(* IEC 61131-3 sources: s7-to-codesys/src/DUTs/S7Compat, 2 files *)

(* ---- ST_S5Counter.dut.st ---- *)
// Назначение: состояние счётчика S5 (слово счётчика C n S7-300/400) для кода, сконвертированного s7conv из
//             STL: CU, CD, установка S, сброс R, разрешение FR, опрос A C, L C, LC C. Значение 0…999; у
//             каждой инструкции, работающей по фронту RLO, своя память фронта. Состояния лежат в
//             генерируемом GVL_S5Counters (массив aCounter, индекс — номер счётчика).
// Автор:      kr0nsch
// Версия:     1.2.0
// Документ:   docs/MAPPING_STL.md, правило s5.counter
TYPE ST_S5Counter :
STRUCT
    iValue : INT;       // значение счётчика, 0…999
    xRloUp : BOOL;      // RLO последней инструкции CU — память фронта
    xRloDown : BOOL;    // RLO последней инструкции CD — память фронта
    xRloSet : BOOL;     // RLO последней инструкции S — память фронта
    xRloFree : BOOL;    // RLO последней инструкции FR — память фронта разрешения
END_STRUCT
END_TYPE

(* ---- ST_S5Timer.dut.st ---- *)
// Назначение: состояние таймера S5 (слово таймера T n S7-300/400) для кода, сконвертированного s7conv из STL:
//             пуск SP, SE, SD, SS, SF, разрешение FR, сброс R, опрос A T, L T, LC T. В S7 таймер — глобальный
//             объект CPU, поэтому состояния лежат в генерируемом GVL_S5Timers (массив aTimer, индекс — номер
//             таймера), а инструкции — функции F_S5* с VAR_IN_OUT. Время — F_S7Now(): в работе TIME(), в
//             тестах — моделируемые часы GVL_S7Clock. Остаток пересчитывается при каждом обращении к таймеру
//             (в S7 его уменьшает часовой процесс CPU асинхронно циклу).
// Автор:      kr0nsch
// Версия:     1.2.0
// Документ:   docs/MAPPING_STL.md, правило s5.timebase; docs/ASSUMPTIONS.md, записи L13–L16
TYPE ST_S5Timer :
STRUCT
    xRunning : BOOL;    // таймер идёт
    xQ : BOOL;          // состояние таймера (опрос A T n)
    xRloStart : BOOL;   // RLO последней инструкции пуска — память фронта пуска (FR её сбрасывает)
    xRloFree : BOOL;    // RLO последней инструкции FR — память фронта разрешения
    xQAtEnd : BOOL;     // состояние по истечении времени: TRUE — SD, SS; FALSE — SP, SE, SF
    tStart : TIME;      // момент пуска (F_S7Now)
    tPreset : TIME;     // заданное время: значение × шкала
    tRest : TIME;       // остаток времени (у остановленного таймера — на момент остановки)
    wBase : WORD;       // шкала времени: 0 — 10 мс, 1 — 100 мс, 2 — 1 с, 3 — 10 с
END_STRUCT
END_TYPE
